# EPICS autosave request: ioc/autoSaveRestore/energy_meter_two_heads.req
file "head.req",	head=$(HEAD1)
file "head.req",	head=$(HEAD2)
